                      Waypoint spat_L_up: motionParameters(blendRadius=0.05); TCP in base x=247.136 y=-17.665 z=397.131 mm, rx=0 ry=-0.0005 rz=3.1068 rad; joints [28.565, -53.55, -103.607, -112.824, 90.132, 120.503] deg
                    MoveJ speed 60 deg/s, acceleration 80 deg/s^2 (useActiveTCP=true optimoveEnabled=false optiMoveSpeed=0.3 optiMoveAcceleration=0.09) feature=Base
                      Waypoint Spatula_otw: TCP in base x=-38.472 y=-263.141 z=425.351 mm, rx=-0.0004 ry=-0.0001 rz=3.0344 rad; joints [-68.119, -57.773, -97.702, -114.504, 90.127, 27.957] deg
                  ElseIf spatula ≟"spatula_M"
                    MoveJ speed 60 deg/s, acceleration 80 deg/s^2 (useActiveTCP=true optimoveEnabled=false optiMoveSpeed=0.3 optiMoveAcceleration=0.09) feature=Base
                      Waypoint Spatula_otw: TCP in base x=-38.472 y=-263.141 z=425.351 mm, rx=-0.0004 ry=-0.0001 rz=3.0344 rad; joints [-68.119, -57.773, -97.702, -114.504, 90.127, 27.957] deg
                      Waypoint spat_M_up: motionParameters(blendRadius=0.05); TCP in base x=245.496 y=-112.113 z=420.344 mm, rx=0 ry=-0.0005 rz=3.0677 rad; joints [5.167, -58.065, -98.393, -113.528, 90.127, 99.337] deg
                    MoveL speed 250 mm/s, acceleration 1200 mm/s^2 (useActiveTCP=true optimoveEnabled=false optiMoveSpeed=0.3 optiMoveAcceleration=0.09) feature=Base
                      Waypoint spat_M_pick: TCP in base x=244.674 y=-111.985 z=192.299 mm, rx=0 ry=-0.0005 rz=3.0677 rad; joints [5.062, -53.127, -134.29, -82.569, 90.166, 99.363] deg
                      URCap Gripper (Robotiq_Grippers, Robotiq Inc.) dataModel(position=100.0, force=30.0, speed=0.0, positionInDouble=100.0, forceInDouble=30.0, speedInDouble=0.0, slaveIds=[9], blocking=true)
                      Waypoint spat_M_up: motionParameters(blendRadius=0.05); TCP in base x=245.496 y=-112.113 z=420.344 mm, rx=0 ry=-0.0005 rz=3.0677 rad; joints [5.167, -58.065, -98.393, -113.528, 90.127, 99.337] deg
                      Waypoint Spatula_otw: TCP in base x=-38.472 y=-263.141 z=425.351 mm, rx=-0.0004 ry=-0.0001 rz=3.0344 rad; joints [-68.119, -57.773, -97.702, -114.504, 90.127, 27.957] deg
                    switch_spat_M := False
                  ElseIf spatula≟"spatula_S"
                    MoveJ speed 60 deg/s, acceleration 80 deg/s^2 (useActiveTCP=true optimoveEnabled=false optiMoveSpeed=0.3 optiMoveAcceleration=0.09) feature=Base
                      Waypoint Spatula_otw: TCP in base x=-38.472 y=-263.141 z=425.351 mm, rx=-0.0004 ry=-0.0001 rz=3.0344 rad; joints [-68.119, -57.773, -97.702, -114.504, 90.127, 27.957] deg
                      Waypoint spat_S_Up_7: motionParameters(blendRadius=0.05); TCP in base x=252.088 y=-159.242 z=423.282 mm, rx=0 ry=-0.0005 rz=3.0677 rad; joints [-5.618, -62.24, -96.192, -111.556, 90.127, 88.551] deg
                    MoveL speed 250 mm/s, acceleration 1200 mm/s^2 (useActiveTCP=true optimoveEnabled=false optiMoveSpeed=0.3 optiMoveAcceleration=0.09) feature=Base
                      Waypoint spat_S_Pick_4: TCP in base x=245.377 y=-158.668 z=192.286 mm, rx=0 ry=-0.0005 rz=3.0677 rad; joints [-5.78, -57.937, -132.467, -79.585, 90.161, 88.525] deg
                      URCap Gripper (Robotiq_Grippers, Robotiq Inc.) dataModel(position=100.0, force=30.0, speed=0.0, positionInDouble=100.0, forceInDouble=30.0, speedInDouble=0.0, slaveIds=[9], blocking=true)
                      Waypoint spat_S_Up_8: motionParameters(blendRadius=0.05); TCP in base x=252.088 y=-159.242 z=423.282 mm, rx=0 ry=-0.0005 rz=3.0677 rad; joints [-5.618, -62.24, -96.192, -111.556, 90.127, 88.551] deg
                      Waypoint Spatula_otw: TCP in base x=-38.472 y=-263.141 z=425.351 mm, rx=-0.0004 ry=-0.0001 rz=3.0344 rad; joints [-68.119, -57.773, -97.702, -114.504, 90.127, 27.957] deg
                    switch_spat_S := False
                  ElseIf spatula≟"spatula_flat_M"
                    MoveJ speed 60 deg/s, acceleration 80 deg/s^2 (useActiveTCP=true optimoveEnabled=false optiMoveSpeed=0.3 optiMoveAcceleration=0.09) feature=Base
                      Waypoint Spatula_otw: TCP in base x=-38.472 y=-263.141 z=425.351 mm, rx=-0.0004 ry=-0.0001 rz=3.0344 rad; joints [-68.119, -57.773, -97.702, -114.504, 90.127, 27.957] deg
                      Waypoint spat_flatM_up: motionParameters(blendRadius=0.05); TCP in base x=229.023 y=-211.443 z=418.634 mm, rx=0 ry=-0.0005 rz=3.0677 rad; joints [-17.294, -63.925, -96.117, -109.949, 90.128, 76.878] deg
                    MoveL speed 250 mm/s, acceleration 1200 mm/s^2 (useActiveTCP=true optimoveEnabled=false optiMoveSpeed=0.3 optiMoveAcceleration=0.09) feature=Base
                      Waypoint spat_flatM_pick: TCP in base x=241.029 y=-208.057 z=192.271 mm, rx=0 ry=-0.0005 rz=3.0677 rad; joints [-16.075, -63.047, -130.143, -76.801, 90.154, 78.231] deg
                      URCap Gripper (Robotiq_Grippers, Robotiq Inc.) dataModel(position=100.0, force=30.0, speed=0.0, positionInDouble=100.0, forceInDouble=30.0, speedInDouble=0.0, slaveIds=[9], blocking=true, robotCompliant=false)
                      Waypoint spat_flatM_up: motionParameters(blendRadius=0.05); TCP in base x=229.023 y=-211.443 z=418.634 mm, rx=0 ry=-0.0005 rz=3.0677 rad; joints [-17.294, -63.925, -96.117, -109.949, 90.128, 76.878] deg
                      Waypoint Spatula_otw: TCP in base x=-38.472 y=-263.141 z=425.351 mm, rx=-0.0004 ry=-0.0001 rz=3.0344 rad; joints [-68.119, -57.773, -97.702, -114.504, 90.127, 27.957] deg
                    switch_spat_F_M := False
                  ElseIf spatula≟"spatula_flat_S"
                    MoveJ speed 60 deg/s, acceleration 80 deg/s^2 (useActiveTCP=true optimoveEnabled=false optiMoveSpeed=0.3 optiMoveAcceleration=0.09) feature=Base
                      Waypoint Spatula_otw: TCP in base x=-38.472 y=-263.141 z=425.351 mm, rx=-0.0004 ry=-0.0001 rz=3.0344 rad; joints [-68.119, -57.773, -97.702, -114.504, 90.127, 27.957] deg
                      Waypoint spat_flatS_up: motionParameters(blendRadius=0.05); TCP in base x=237.652 y=-253.944 z=403.961 mm, rx=0 ry=-0.0005 rz=3.0677 rad; joints [-24.273, -68.411, -95.947, -105.635, 90.132, 69.906] deg
                    MoveL speed 250 mm/s, acceleration 1200 mm/s^2 (useActiveTCP=true optimoveEnabled=false optiMoveSpeed=0.3 optiMoveAcceleration=0.09) feature=Base
                      Waypoint spat_flatS_pick: TCP in base x=241.326 y=-251.726 z=192.257 mm, rx=0 ry=-0.0005 rz=3.0677 rad; joints [-23.749, -68.568, -127.154, -74.27, 90.149, 70.556] deg
                      URCap Gripper (Robotiq_Grippers, Robotiq Inc.) dataModel(position=100.0, force=30.0, speed=0.0, positionInDouble=100.0, forceInDouble=30.0, speedInDouble=0.0, slaveIds=[9], blocking=true, robotCompliant=false)
                      Waypoint spat_flatS_up: motionParameters(blendRadius=0.05); TCP in base x=237.652 y=-253.944 z=403.961 mm, rx=0 ry=-0.0005 rz=3.0677 rad; joints [-24.273, -68.411, -95.947, -105.635, 90.132, 69.906] deg
                      Waypoint Spatula_otw: TCP in base x=-38.472 y=-263.141 z=425.351 mm, rx=-0.0004 ry=-0.0001 rz=3.0344 rad; joints [-68.119, -57.773, -97.702, -114.504, 90.127, 27.957] deg
                    switch_spat_F_S := False
                  weight_value := get_weight()
                  Script: auto_tilt_and_scoop(W_now, target_weight, weight_value)
                URCap Approach Pose (SensoPart VISOR Robotic, SensoPart Industriesensorik GmbH) dataModel(visorJointSpeed=10.0, visorJointAcc=15.0, visorOffsetZ=-30.0); state(isChildrenLocked=true)
                URCap Target Pose (SensoPart VISOR Robotic, SensoPart Industriesensorik GmbH) dataModel(visorToolSpeed=20.0, visorToolAcc=50.0); state(isChildrenLocked=true)
                Folder Close Gripper
                  dispense_pos := get_actual_tcp_pose()
                  Loop While (checkContinuously=true) expression=weight_value≤target_weight
                    MoveL speed 250 mm/s, acceleration 1200 mm/s^2 (useActiveTCP=true optimoveEnabled=false optiMoveSpeed=0.3 optiMoveAcceleration=0.09) feature=Base
                      Waypoint Variable (Variable): motionParameters(jointSpeed=0.436332 jointAcceleration=0.523599 cartesianSpeed=0.1 cartesianAcceleration=0.2); variable=dispense_pos
                      Script: log_weight()
                      Wait Sleep waitTime=0.5
                      If level≥90.0
                        Script: Rotate()
                      If level≤85
                        Script: tilt_to_home()
                      Wait Sleep waitTime=0.5
                      Start_thread := True
                      vib_thread := True
                      SuppressedNode
                        tilt_angle := current_pose[5]
                      Wait Sleep waitTime=0.5
                      SuppressedNode
                        Loop While (checkContinuously=true) expression=diff>3.0
                          tilt_pose := pose_trans(get_actual_tcp_pose(), p[0, 0, 0, 0, 0, 1.0])
                          Script: movel(tilt_pose, a=0.1, v=0.1, r=0.00001)
                          tilt_pose := pose_trans(get_actual_tcp_pose(), p[0, 0, 0, 0, 0, -1.0])
                          Script: movel(tilt_pose, a=0.1, v=0.1, r=0.00001)
                      If diff ≥(target_g +(0.1*target_g))
                        tilt_pose := pose_trans(get_actual_tcp_pose(), p[0, 0, 0, 0, 0, 2.0])
                        Script: movel(tilt_pose, a=0.1, v=0.1, r=0.00001)
                      Else 
                        Loop While (checkContinuously=true) expression=weight_value≤target_weight and tilt_angle≥(-1.999) and tilt_angle≤0.5
                          current_error := target_weight-weight_value
                          Integral_error := Integral_error+current_error*dt
                          derivative := (current_error-previous_error)/dt
                          tilt_increment := (kp*current_error)+(ki*Integral_error)+(kd*derivative)
                          current_pose := get_actual_tcp_pose()
                          tilt_angle := current_pose[5]
                          tilt_pose := pose_trans(current_pose, p[0, 0, 0, 0, 0, tilt_increment])
                          Script: movel(tilt_pose, a=0.1, v=0.1, r=0.00001)
                          previous_error := current_error
                      Start_thread := False
                      SuppressedNode
                        Waypoint Waypoint_64: motionParameters(jointSpeed=1.047198 jointAcceleration=1.396263 cartesianSpeed=0.03 cartesianAcceleration=0.1 blendRadius=0.05); TCP in base x=-542.998 y=-117.021 z=221.977 mm, rx=1.8981 ry=-0.7227 rz=1.5827 rad; joints [-123.845, -120.87, -101.018, -172.406, 14.907, 127.864] deg
                      weight_value := get_weight()
                      tilt_angle := -1
                      Wait Sleep waitTime=0.5
                      vib_thread := False
                      MoveL speed 250 mm/s, acceleration 500 mm/s^2 (useActiveTCP=true optimoveEnabled=false optiMoveSpeed=0.3 optiMoveAcceleration=0.09) feature=Base
                        Waypoint Variable (Variable): variable=dispense_pos
                      Script: compute_level_percent(W_now, weight_value)
                      Script: send_level_info()
                      Script: spatula = select_spatula(Pow_name, level, diff)
                      Wait Sleep waitTime=0.2
                      SuppressedNode
                        Script: spatula = str_cat("", spatula)
                      Integral_error := 0
                      current_error := 0
                      previous_error := 0
                      Set AnalogOutput pin=analog_out[0]; analogValue=0
                      Wait Sleep waitTime=0.2
                      Script: send_spatula_info()
                      If spatula ≟ "spatula_M" and switch_spat_M≟ True
                        MoveJ speed 60 deg/s, acceleration 80 deg/s^2 (useActiveTCP=true optimoveEnabled=false optiMoveSpeed=0.3 optiMoveAcceleration=0.09) feature=Base
                          Waypoint Spatula_otw: TCP in base x=-38.472 y=-263.141 z=425.351 mm, rx=-0.0004 ry=-0.0001 rz=3.0344 rad; joints [-68.119, -57.773, -97.702, -114.504, 90.127, 27.957] deg
                          Waypoint spat_L_up: TCP in base x=247.136 y=-17.665 z=397.131 mm, rx=0 ry=-0.0005 rz=3.1068 rad; joints [28.565, -53.55, -103.607, -112.824, 90.132, 120.503] deg
                        MoveL speed 250 mm/s, acceleration 1200 mm/s^2 (useActiveTCP=true optimoveEnabled=false optiMoveSpeed=0.3 optiMoveAcceleration=0.09) feature=Base
                          Waypoint spat_L_side: TCP in base x=247.134 y=-17.634 z=289.063 mm, rx=0 ry=-0.0005 rz=3.1068 rad; joints [28.487, -49.174, -121.365, -99.443, 90.16, 120.484] deg
                          Waypoint spat_L_lift: TCP in base x=245.402 y=-67.432 z=289.049 mm, rx=0 ry=-0.0005 rz=3.1068 rad; joints [16.24, -50.411, -121.005, -98.568, 90.16, 108.238] deg
                          Waypoint spat_L_pick: TCP in base x=242.469 y=-67.302 z=193.171 mm, rx=0 ry=-0.0005 rz=3.1068 rad; joints [16.429, -49.275, -135.385, -85.324, 90.17, 108.483] deg
                          URCap Gripper (Robotiq_Grippers, Robotiq Inc.) dataModel(position=0.0, force=30.0, speed=100.0, positionInDouble=0.0, forceInDouble=30.0, speedInDouble=100.0, slaveIds=[9], blocking=true)
                          Waypoint spat_M_pick: TCP in base x=244.674 y=-111.985 z=192.299 mm, rx=0 ry=-0.0005 rz=3.0677 rad; joints [5.062, -53.127, -134.29, -82.569, 90.166, 99.363] deg
                          URCap Gripper (Robotiq_Grippers, Robotiq Inc.) dataModel(position=100.0, force=30.0, speed=0.0, positionInDouble=100.0, forceInDouble=30.0, speedInDouble=0.0, slaveIds=[9], blocking=true)
                          Waypoint spat_M_up: TCP in base x=245.496 y=-112.113 z=420.344 mm, rx=0 ry=-0.0005 rz=3.0677 rad; joints [5.167, -58.065, -98.393, -113.528, 90.127, 99.337] deg
                          Waypoint Spatula_otw: TCP in base x=-38.472 y=-263.141 z=425.351 mm, rx=-0.0004 ry=-0.0001 rz=3.0344 rad; joints [-68.119, -57.773, -97.702, -114.504, 90.127, 27.957] deg
                        switch_spat_M := False
                      ElseIf spatula ≟ "spatula_S" and switch_spat_S ≟ True
                        MoveL speed 250 mm/s, acceleration 1200 mm/s^2 (useActiveTCP=true optimoveEnabled=false optiMoveSpeed=0.3 optiMoveAcceleration=0.09) feature=Base
                          Waypoint Spatula_otw: TCP in base x=-38.472 y=-263.141 z=425.351 mm, rx=-0.0004 ry=-0.0001 rz=3.0344 rad; joints [-68.119, -57.773, -97.702, -114.504, 90.127, 27.957] deg
                          Waypoint spat_M_up: TCP in base x=245.496 y=-112.113 z=420.344 mm, rx=0 ry=-0.0005 rz=3.0677 rad; joints [5.167, -58.065, -98.393, -113.528, 90.127, 99.337] deg
                          Waypoint spat_M_pick: TCP in base x=244.674 y=-111.985 z=192.299 mm, rx=0 ry=-0.0005 rz=3.0677 rad; joints [5.062, -53.127, -134.29, -82.569, 90.166, 99.363] deg
                          URCap Gripper (Robotiq_Grippers, Robotiq Inc.) dataModel(position=0.0, force=30.19607843137255, speed=100.0, positionInDouble=0.0, forceInDouble=30.19607843137255, speedInDouble=100.0, slaveIds=[9], blocking=true)
                          Waypoint spat_S_pick: TCP in base x=238.159 y=-157.927 z=192.632 mm, rx=0 ry=-0.0005 rz=3.0677 rad; joints [-5.778, -56.616, -132.95, -80.422, 90.162, 88.526] deg
                          URCap Gripper (Robotiq_Grippers, Robotiq Inc.) dataModel(position=100.0, force=30.19607843137255, speed=0.0, positionInDouble=100.0, forceInDouble=30.19607843137255, speedInDouble=0.0, slaveIds=[9], blocking=true)
                          Waypoint spat_S_up: TCP in base x=244.261 y=-164.467 z=417.088 mm, rx=0 ry=-0.0005 rz=3.0677 rad; joints [-6.934, -61.411, -97.537, -111.041, 90.129, 87.239] deg
                          Waypoint Spatula_otw: TCP in base x=-38.472 y=-263.141 z=425.351 mm, rx=-0.0004 ry=-0.0001 rz=3.0344 rad; joints [-68.119, -57.773, -97.702, -114.504, 90.127, 27.957] deg
                        switch_spat_S := False
                      ElseIf spatula≟"spatula_flat_S"  and switch_spat_F_S ≟ True
                        MoveL speed 250 mm/s, acceleration 1200 mm/s^2 (useActiveTCP=true optimoveEnabled=false optiMoveSpeed=0.3 optiMoveAcceleration=0.09) feature=Base
                          Waypoint Spatula_otw: TCP in base x=-38.472 y=-263.141 z=425.351 mm, rx=-0.0004 ry=-0.0001 rz=3.0344 rad; joints [-68.119, -57.773, -97.702, -114.504, 90.127, 27.957] deg
                          Waypoint spat_flatM_up: TCP in base x=229.023 y=-211.443 z=418.634 mm, rx=0 ry=-0.0005 rz=3.0677 rad; joints [-17.294, -63.925, -96.117, -109.949, 90.128, 76.878] deg
                          Waypoint spat_flatM_pick: TCP in base x=241.029 y=-208.057 z=192.271 mm, rx=0 ry=-0.0005 rz=3.0677 rad; joints [-16.075, -63.047, -130.143, -76.801, 90.154, 78.231] deg
                          URCap Gripper (Robotiq_Grippers, Robotiq Inc.) dataModel(position=0.0, force=30.0, speed=0.0, positionInDouble=0.0, forceInDouble=30.0, speedInDouble=0.0, slaveIds=[9], blocking=true, robotCompliant=false)
                          Waypoint spat_flatS_pick: TCP in base x=241.326 y=-251.726 z=192.257 mm, rx=0 ry=-0.0005 rz=3.0677 rad; joints [-23.749, -68.568, -127.154, -74.27, 90.149, 70.556] deg
                          URCap Gripper (Robotiq_Grippers, Robotiq Inc.) dataModel(position=100.0, force=30.0, speed=0.0, positionInDouble=100.0, forceInDouble=30.0, speedInDouble=0.0, slaveIds=[9], blocking=true, robotCompliant=false)
                          Waypoint spat_flatS_up: TCP in base x=237.652 y=-253.944 z=403.961 mm, rx=0 ry=-0.0005 rz=3.0677 rad; joints [-24.273, -68.411, -95.947, -105.635, 90.132, 69.906] deg
                          Waypoint Spatula_otw: TCP in base x=-38.472 y=-263.141 z=425.351 mm, rx=-0.0004 ry=-0.0001 rz=3.0344 rad; joints [-68.119, -57.773, -97.702, -114.504, 90.127, 27.957] deg
                        switch_spat_F_S := False
                      Script: auto_tilt_and_scoop(W_now, target_weight, weight_value)
                      Wait Sleep waitTime=0.5
                  Start_thread := False
                  Wait Sleep waitTime=0.5
                  vib_thread := False
                  SuppressedNode
                    Script: Rotate()
                URCap Exit Pose (SensoPart VISOR Robotic, SensoPart Industriesensorik GmbH) dataModel(visorOffsetZ=0.0); state(isChildrenLocked=true)
              URCap No Object Detected (SensoPart VISOR Robotic, SensoPart Industriesensorik GmbH) dataModel(Variable(key=visorNoObjCountVar, variable=easyPickNoObj_4))
                Popup Message (haltProgram=false message=No weigh scale detected inputType=Text)
          SuppressedNode
            Task := "Dosing"
          SuppressedNode
            Script: scooping_init()
          MoveJ speed 60 deg/s, acceleration 80 deg/s^2 (useActiveTCP=true optimoveEnabled=false optiMoveSpeed=0.3 optiMoveAcceleration=0.09) feature=Base
            Waypoint Variable (Variable): motionParameters(jointSpeed=0.436332 jointAcceleration=0.523599 cartesianSpeed=0.1 cartesianAcceleration=0.2); variable=dispense_pos
          Script: after_scoop()
          SuppressedNode
            Folder powder dispensing
              SuppressedNode
                Target_weight := Target_weight/1000
              Loop While (checkContinuously=false) expression=Weight_value<Target_weight
                Script: auto_tilt_and_scoop(W_now, Target_weight, Weight_value)
                Start_thread := True
                MoveL speed 250 mm/s, acceleration 1200 mm/s^2 (useActiveTCP=true optimoveEnabled=false optiMoveSpeed=0.3 optiMoveAcceleration=0.09) feature=Base
                  Waypoint Variable (Variable): motionParameters(jointSpeed=0.436332 jointAcceleration=0.523599 cartesianSpeed=0.05 cartesianAcceleration=0.2); variable=dispense_pos
                  Wait Sleep waitTime=0.5
                  Script: Rotate()
                  Wait Sleep waitTime=0.5
                MoveL speed 250 mm/s, acceleration 1200 mm/s^2 (useActiveTCP=true optimoveEnabled=false optiMoveSpeed=0.3 optiMoveAcceleration=0.09) feature=Base
                  Start_thread := True
                  vib_mot_thread := True
                  tilt_angle := current_pose[5]
                  Wait Sleep waitTime=0.5
                  SuppressedNode
                    Loop While (checkContinuously=true) expression=diff>3.0
                      tilt_pose := pose_trans(get_actual_tcp_pose(), p[0, 0, 0, 0, 0, 1.0])
                      Script: movel(tilt_pose, a=0.1, v=0.1, r=0.00001)
                      tilt_pose := pose_trans(get_actual_tcp_pose(), p[0, 0, 0, 0, 0, -1.0])
                      Script: movel(tilt_pose, a=0.1, v=0.1, r=0.00001)
                  If diff>3.0
                    tilt_pose := pose_trans(get_actual_tcp_pose(), p[0, 0, 0, 0, 0, 2.0])
                    Script: movel(tilt_pose, a=0.1, v=0.1, r=0.00001)
                  ElseIf diff≤3.0
                    Loop While (checkContinuously=false) expression=Weight_value≤Target_weight and tilt_angle≥(-1.999) and tilt_angle≤0
                      current_error := Target_weight-Weight_value
                      Integral_error := Integral_error+current_error*dt
                      derivative := (current_error-previous_error)/dt
                      tilt_increment := (kp*current_error)+(ki*Integral_error)+(kd*derivative)
                      current_pose := get_actual_tcp_pose()
                      tilt_angle := current_pose[5]
                      tilt_pose := pose_trans(current_pose, p[0, 0, 0, 0, 0, tilt_increment])
                      Script: movel(tilt_pose, a=0.1, v=0.1, r=0.00001)
                      previous_error := current_error
                  Start_thread := False
                  SuppressedNode
                    Waypoint Waypoint_64: motionParameters(jointSpeed=1.047198 jointAcceleration=1.396263 cartesianSpeed=0.03 cartesianAcceleration=0.1 blendRadius=0.05); TCP in base x=-542.998 y=-117.021 z=221.977 mm, rx=1.8981 ry=-0.7227 rz=1.5827 rad; joints [-123.845, -120.87, -101.018, -172.406, 14.907, 127.864] deg
                  Weight_value := get_weight()
                  Wait Sleep waitTime=0.5
                  tilt_angle := -1
                  vib_mot_thread := False
                  MoveL speed 50 mm/s, acceleration 300 mm/s^2 (useActiveTCP=true optimoveEnabled=false optiMoveSpeed=0.3 optiMoveAcceleration=0.09) feature=Base
                    Waypoint Variable (Variable): motionParameters(jointSpeed=0.436332 jointAcceleration=0.523599 cartesianSpeed=0.05 cartesianAcceleration=0.2); variable=dispense_pos
                  Integral_error := 0
                  current_error := 0
                  previous_error := 0
                  Set AnalogOutput pin=analog_out[0]; analogValue=0
                Script: movel(pose_trans(dispense_pos, p[-0.02,0,0,0,0,0]))
              SuppressedNode
                MoveL speed 250 mm/s, acceleration 1200 mm/s^2 (useActiveTCP=true optimoveEnabled=false optiMoveSpeed=0.3 optiMoveAcceleration=0.09) feature=Base
                  Waypoint aftr_scoo3: motionParameters(jointSpeed=1.047198 jointAcceleration=1.396263 cartesianSpeed=0.1 cartesianAcceleration=0.3); TCP in base x=-289.76 y=-315.385 z=303.744 mm, rx=0.16 ry=1.6274 rz=-0.3449 rad; joints [-76.632, -96.313, -113.776, -155.476, 32.027, -78.1] deg
                  Waypoint ftr_scoop2: motionParameters(jointSpeed=1.047198 jointAcceleration=1.396263 cartesianSpeed=0.1 cartesianAcceleration=0.4); TCP in base x=194.287 y=-495.78 z=282.072 mm, rx=-0.179 ry=1.6121 rz=-0.016 rad; joints [-34.133, -129.723, -68.393, -165.549, 50.138, -80.843] deg
                  Waypoint aftr_scoop1: motionParameters(jointSpeed=1.047198 jointAcceleration=1.396263 cartesianSpeed=0.1 cartesianAcceleration=0.4); TCP in base x=138.504 y=-514.48 z=214.154 mm, rx=-0.1348 ry=1.5599 rz=-0.0592 rad; joints [-39.422, -130.004, -76.262, -153.157, 47.788, -83.41] deg
                  Waypoint After_disp_3: motionParameters(jointSpeed=1.047198 jointAcceleration=1.396263 cartesianSpeed=0.1 cartesianAcceleration=0.4); TCP in base x=125.935 y=-585.611 z=299.546 mm, rx=0.9596 ry=-0.1344 rz=2.8807 rad; joints [-54.056, -115.535, -63.235, -120.118, 65.773, 48.319] deg
                  Set AnalogOutput pin=analog_out[0]; analogValue=3
                  Wait Sleep waitTime=2
                  Set AnalogOutput pin=analog_out[0]; analogValue=0
                  Waypoint aftr_scoop1: TCP in base x=138.504 y=-514.48 z=214.154 mm, rx=-0.1348 ry=1.5599 rz=-0.0592 rad; joints [-39.422, -130.004, -76.262, -153.157, 47.788, -83.41] deg
                  Waypoint ftr_scoop2: motionParameters(jointSpeed=1.047198 jointAcceleration=1.396263 cartesianSpeed=0.1 cartesianAcceleration=0.4); TCP in base x=194.287 y=-495.78 z=282.072 mm, rx=-0.179 ry=1.6121 rz=-0.016 rad; joints [-34.133, -129.723, -68.393, -165.549, 50.138, -80.843] deg
                  Waypoint Waypoint_63: motionParameters(blendRadius=0.05); TCP in base x=101.295 y=-465.376 z=381.756 mm, rx=0.9726 ry=-0.1584 rz=2.8872 rad; joints [-48.863, -99.659, -71.872, -130.079, 68.56, 52.636] deg; TCP offset x=0 y=0 z=161 mm, rx=3.1415 ry=0 rz=0 rad
                  Waypoint Start: motionParameters(jointSpeed=1.047198 jointAcceleration=1.396263 cartesianSpeed=0.15 cartesianAcceleration=0.6); TCP in base x=-33.065 y=-365.399 z=389.873 mm, rx=0 ry=0 rz=2.7258 rad; joints [-73.774, -70.638, -96.716, -102.629, 90.121, 40.001] deg; TCP offset x=0 y=0 z=161 mm, rx=3.1415 ry=0 rz=0 rad
                  Popup Message (haltProgram=false message=Powder dispensed successfully... inputType=Text)
              SuppressedNode
                Script: tilt()
          SuppressedNode
            Script: tilt_send()
      Case (caseValue=44)
        Folder Decap Container for recipe [hidden by the author, left out]
      Case (caseValue=45)
        Folder Place the decapped container- recipe [hidden by the author, left out]
      Case (caseValue=46)
        Folder Powder dosing for recipe [hidden by the author, left out]
      Case (caseValue=47)
        Folder Pick containers [hidden by the author, left out]
      Case (caseValue=48)
        Folder QR detections [hidden by the author, left out]
  SuppressedNode
    '=========='
  SuppressedNode
    Folder PostSettings [hidden by the author, left out]
